// TIA Portal V20 export
// export: Created 2026-10-12T04:58:21.0883789Z, ExportSetting WithDefaults, DisplayName Totally Integrated Automation Portal, DisplayVersion V20, DisplayName TIA Portal Openness, DisplayVersion V20, DisplayName TIA Portal Teamcenter Gateway, DisplayVersion V20, DisplayName TIA Portal Version Control Interface, DisplayVersion V20, DisplayName SINAMICS Startdrive Advanced, DisplayVersion V20 SP1 Update 2, DisplayName SINAMICS Startdrive G110M, G120, G120C, G120D, G120P, G115D, DisplayVersion V20 SP1 Update 2, DisplayName SINAMICS Startdrive G130, G150, S120, S150, SINAMICS MV, G220, S200, S210, DisplayVersion V20 SP1 Update 2, DisplayName STEP 7 Professional, DisplayVersion V20, DisplayName STEP 7 Safety, DisplayVersion V20, DisplayName WinCC Basic/Comfort/Advanced, DisplayVersion V20, DisplayName WinCC Professional, DisplayVersion V20, DisplayName WinCC Unified, DisplayVersion V20
FUNCTION "FRK_DecisionClear" : Void   // FC88, SCL
{ S7_Optimized_Access := 'TRUE' }
VERSION : 0.1
// stored: AutoNumber true, IsIECCheckEnabled false, SetENOAutomatically false, UDAEnableTagReadback false
   VAR_IN_OUT
      Slot : "FRK_DecisionSlot";
   END_VAR
   VAR_TEMP
      Index : Int;
   END_VAR
BEGIN

   #Slot.Request.Prompt := WSTRING#'';
   #Slot.Request.SourcePath := WSTRING#'';
   #Slot.Request.Default := 0;
   #Slot.Request.Timeout := T#0ms;
   FOR #Index := 1 TO 6 DO
       #Slot.Request.Options[#Index] := '';
   END_FOR;
   #Slot.Answer := 0;
   #Slot.Owner := 0;
   #Slot.OverlapLogged := FALSE;
   #Slot.ResolutionLogged := FALSE;
END_FUNCTION
